{attribute 'no_assign'}
FUNCTION_BLOCK FB_LN_WTURBINE_LD0_WGEN1 EXTENDS FB_AcsiCommonLogicalNodeClass
VAR_INPUT
	Beh: FB_DO_WTURBINE_LD0_WGEN1_Beh := (sClass:='ENS', bLinkResult:=THIS^.AddDataToContainer(ipData:=Beh));
	RotSpd: FB_DO_WTURBINE_LD0_WGEN1_RotSpd := (sClass:='MV', bLinkResult:=THIS^.AddDataToContainer(ipData:=RotSpd));
END_VAR
VAR
END_VAR

END_FUNCTION_BLOCK

(* stored: Version 1.1.0.1
   POU FB_LN_WTURBINE_LD0_WGEN1: Id {da2921c2-550f-4c6b-ac13-6d9f6223cb3f}, SpecialFunc None *)
